Universal Robots PolyScope program: Prog_Name_That_Is_Very_Long_123.urp

Program Prog_Name_That_Is_Very_Long_123 (createdIn=3.0.0 lastSavedIn=3.0.0 directory=. installation=default)
Robot Program (runOnlyOnce=true motionType=MoveJ speed=1.047198 acceleration=1.396263 useActiveTCP=false)
  Script file Prog_Name_That_Is_Very_Long_123.script
    | def Prog_Name_That_Is_Very_Long_123():
    |   # Global parameters:
    |   global speed_ms    = 0.250
    |   global speed_rads  = 0.750
    |   global accel_mss   = 1.200
    |   global accel_radss = 1.200
    |   global blend_radius_m = 0.001
    |   global ref_frame = p[0,0,0,0,0,0]
    | 
    |   #
    |   # TO REMOVE HEADER:
    |   # Go to "Program" -> "Post-Processor Editor"
    |   # Select "Universal Robots"
    |   # Set "INCLUDE_HEADER" to "False"
    |   #
    |   #--------------------------
    |   # Add any default subprograms here
    |   # For example, to drive a gripper as a program call:
    |   # def Gripper_Open():
    |   #   ...
    |   # end
    |   #
    |   # Example to drive a spray gun:
    |   def SprayOn(value):
    |     # use the value as an output:
    |     DO_SPRAY = 5
    |     if value == 0:
    |       set_standard_digital_out(DO_SPRAY, False)
    |     else:
    |       set_standard_digital_out(DO_SPRAY, True)
    |     end
    |   end
    | 
    |   # Example to drive an extruder:
    |   def Extruder(value):
    |     # use the value as an output:
    |     if value < 0:
    |       # stop extruder
    |     else:
    |       # start extruder
    |     end
    |   end
    | 
    |   # Example to move an external axis
    |   def MoveAxis(value):
    |     # use the value as an output:
    |     DO_AXIS_1 = 1
    |     DI_AXIS_1 = 1
    |     if value <= 0:
    |       set_standard_digital_out(DO_AXIS_1, False)
    | 
    |       # Wait for digital input to change state
    |       #while (get_standard_digital_in(DI_AXIS_1) != False):
    |       #  sync()
    |       #end
    |     else:
    |       set_standard_digital_out(DO_AXIS_1, True)
    | 
    |       # Wait for digital input to change state
    |       #while (get_standard_digital_in(DI_AXIS_1) != True):
    |       #  sync()
    |       #end
    |     end
    |   end
    |   #--------------------------
    | 
    | 
    |   # Main program:
    |   # Program generated by VerticalBot Studio for UR5e on 25/10/2026 12:00:00
    |   # Using nominal kinematics.
    |   ref_frame = p[0.000000, 0.000000, 0.000000, 0.000000, 0.000000, 0.000000]
    |   set_tcp(p[0.010000, 0.000000, 0.120000, 0.000000, 0.261799, 0.000000])
    |   speed_ms    = 1.000
    |   blend_radius_m = 0.010
    |   movej([-0.523599, -1.745329, 1.570796, -1.396263, -1.570796, 0.349066],accel_radss,speed_rads,0,0.010)
    |   movel(pose_trans(ref_frame,p[-0.421760, 0.353029, 0.380392, 3.048452, 0.496356, 0.454618]),accel_mss,speed_ms,0,0.010)
    |   blend_radius_m = 0.001
    |   movel(pose_trans(ref_frame,p[-0.384494, 0.350433, 0.368074, 3.036811, 0.389569, 0.461666]),accel_mss,speed_ms,0,0.001)
    |   halt() # reimplement this function to force stop
    |   sleep(1.500)
    |   popup("Say "hi" to the operator","Message",False,False,blocking=False)
    |   # A long comment line that exceeds the usual controller limits for comments by far, really
    |   set_tool_digital_out(2, False)
    |   OUT_A = 1
    |   while (get_standard_digital_in(4) != False):
    |     sync()
    |   end
    |   while (IN_B != True):
    |     sync()
    |   end
    |   Program_With_A_Long_Name_ABCDEFGHIJ()
    |   ref_frame = p[0.250000, 0.300000, -0.010000, 0.000000, 0.000000, 1.570796]
    |   set_tcp(p[0.010000, 0.000000, 0.120000, 0.000000, 0.261799, 0.000000])
    |   speed_rads  = 0.524
    |   accel_radss = 1.745
    |   movel(pose_trans(ref_frame,p[-0.421760, 0.353029, 0.380392, 3.048452, 0.496356, 0.454618]),accel_mss,speed_ms,0,0.001)
    |   blend_radius_m = 0.000
    |   movej([-0.523599, -1.745329, 1.570796, -1.396263, -1.570796, 0.349066],accel_radss,speed_rads,0,0.000)
    |   # End of main program
    | end
    | 
    | Prog_Name_That_Is_Very_Long_123()
